Fanuc KAREL source: KA00029.KL

PROGRAM KA00029
%NOLOCKGROUP
VAR
  SRC: BOOLEAN
  DST: POSITION
BEGIN
  SRC = TRUE
  DST = SRC
END KA00029
